(*
SPDX-FileCopyrightText: © 2026 Oleksandr Tiutyk <trofimich@gmail.com>
SPDX-License-Identifier: MIT
License: https://opensource.org/license/mit
*)

(*!
<summary>Injects a configurable file-manager start preparation exception.</summary>
<description>
Set RefuseStart while READY. With refusal disabled, the probe runs the real file-manager preparation hook.
The test cancels accepted starts before driving native acquisition.
</description>
*)

FUNCTION_BLOCK FileManagerStartRefusalProbe EXTENDS TOF_FileSystem.FileContentManager
VAR_STAT
	_ProbeClassName : STRING := __POUNAME();
END_VAR
VAR_INPUT
	//! <summary>Requests a synthetic preparation exception on the next Start.</summary>
	RefuseStart : BOOL;
END_VAR

(*!
<summary>Raises the requested test exception or delegates to normal file-manager preparation.</summary>
*)
METHOD PROTECTED OnBeforeStart
IF RefuseStart THEN
	TOF_Core.Exceptions.ThrowStandard(
		sourceNamespaceName := NamespaceName,
		sourceClassName := ClassName,
		sourcePOUName := __POUNAME(),
		sourcePosition := __POSITION(),
		message := "Synthetic file-manager Start refusal"
	);
END_IF

SUPER^.OnBeforeStart();
END_METHOD

(*!
<summary>Borrows initialized read-only type metadata without exceptions or resource initialization.</summary>
*)
PROPERTY ClassName : REFERENCE TO STRING
GET
ClassName REF= _ProbeClassName;
END_GET
END_PROPERTY

(*!
<summary>Borrows compiler-initialized read-only metadata identifying the test namespace.</summary>
*)
PROPERTY NamespaceName : REFERENCE TO STRING
GET
NamespaceName REF= CurrentNamespace.Name;
END_GET
END_PROPERTY

(*!
<summary>Reports the size of this concrete probe in bytes.</summary>
*)
PROPERTY SelfSize : ULINT
GET
SelfSize := XSIZEOF(THIS^);
END_GET
END_PROPERTY

END_FUNCTION_BLOCK

(* stored: Version 1.1.0.1
   POU FileManagerStartRefusalProbe: Id {2bf42914-152b-41df-9974-f86511bec283}, SpecialFunc None
   Method OnBeforeStart: Id {f08737f4-ec9a-43a7-8f80-62886edeac76}
   Property ClassName: Id {e8e38f7c-791d-42e0-b6af-bbc729c8944f}
   Get Get: Id {c6235568-2f9e-48a7-9e5f-a2870fcef483}
   Property NamespaceName: Id {1f83b9b2-7697-4e62-9cf2-4a5972664c10}
   Get Get: Id {15ac08c7-b1e6-4d2c-ae63-7500b3f6e6ac}
   Property SelfSize: Id {3d18460c-d2c2-46bc-8ea6-6ac1eb262c04}
   Get Get: Id {bdb9990a-9032-46c0-af4f-60c7d7b5b2d4} *)
